INTERFACE iRoom

METHOD LightsOff
VAR_INPUT
END_VAR
END_METHOD

METHOD LightsOn
VAR_INPUT
END_VAR
END_METHOD

METHOD ShuttersClose
VAR_INPUT
END_VAR
END_METHOD

METHOD ShuttersOpen
VAR_INPUT
END_VAR
END_METHOD

END_INTERFACE

(* stored: Version 1.1.0.1
   Itf iRoom: Id {50cbef3a-567f-429c-942e-dee4c1d64343}
   Method LightsOff: Id {0d1e2a1f-7258-4ee6-ac7a-f11e25a09f6f}
   Method LightsOn: Id {cdc9bfcb-b5cd-47b6-8cc3-8812f8a92317}
   Method ShuttersClose: Id {7866c99d-9838-49be-8223-9db3c85ef106}
   Method ShuttersOpen: Id {e1c9cc61-3b11-4a04-8e31-dd3be03c7065} *)
